(*
SPDX-FileCopyrightText: c 2026 Oleksandr Tiutyk <trofimich@gmail.com>
SPDX-License-Identifier: MIT
License: https://opensource.org/license/mit
*)

(*!
<summary>Checks the native wrapper message in HIDDEN, LOCAL and UTC modes.</summary>
<description>
Uses one task and stays at a stable address while assertions are bound to this instance.
</description>
*)

{attribute 'no_assign'}
{attribute 'no_explicit_call' := 'do not call this function block directly'}
FUNCTION_BLOCK SystemExceptionTimestampFormattingTest EXTENDS TOF_Testing.SingleCycleTest
VAR_STAT
	{attribute 'hide'}
	_ClassName : STRING := __POUNAME();
END_VAR

(*!
<summary>Checks the native wrapper message in HIDDEN, LOCAL and UTC modes.</summary>
<description>
Uses the borrowed wrapper during one callback. The timestamp expectations use the IEC conversion of
captured values and a separately assembled expected message.
</description>
*)
METHOD PROTECTED ExecuteTest
VAR
	exception : TOF_Core.IException;
	hidden : TOF_Core.ERROR_MESSAGE;
	message : TOF_Core.ERROR_MESSAGE;
	expected : WSTRING(255);
	formattingFailed : BOOL;
END_VAR
exception := TOF_Core.ExceptionManager.GetLastException(
	exceptionCode := __SYSTEM.ExceptionCode.RTSEXCPT_ACCESS_VIOLATION,
	catchPointNamespaceName := 'TimestampTest',
	catchPointPOUName := 'NativeCatch',
	catchPointPosition := 'P1'
);

IF exception = 0 THEN
	RecordFailure(message := "The captured native code must provide a wrapper");
	RETURN;
END_IF

hidden := exception.GetMessage(timestampDisplayMode := TOF_Core.TIMESTAMP_DISPLAY_MODE.HIDDEN);
Assert.ThatBool(
	actual := Tc2_Standard.WRIGHT(STR := hidden, SIZE := 31) = "TimestampTest.NativeCatch at P1",
	message := "The hidden timestamp mode must end with the supplied catch location"
).IsTrue();

expected := Tc2_Utilities.WCONCAT(STR1 := hidden, STR2 := " at ");
expected := Tc2_Utilities.WCONCAT(STR1 := expected, STR2 := TO_WSTRING(exception.LocalTimestamp));
formattingFailed := FALSE;

// A formatter exception is recorded for this mode before proceeding to the next check.
__TRY
	message := exception.GetMessage(timestampDisplayMode := TOF_Core.TIMESTAMP_DISPLAY_MODE.LOCAL);
__CATCH
	formattingFailed := TRUE;
__ENDTRY

Assert.ThatBool(
	actual := NOT formattingFailed AND_THEN message = expected,
	message := "LOCAL must append its captured timestamp"
).IsTrue();

expected := Tc2_Utilities.WCONCAT(STR1 := hidden, STR2 := " at ");
expected := Tc2_Utilities.WCONCAT(STR1 := expected, STR2 := TO_WSTRING(exception.UtcTimestamp));
expected := Tc2_Utilities.WCONCAT(STR1 := expected, STR2 := "UTC");
formattingFailed := FALSE;

// A formatter exception is recorded for this mode before proceeding to the next check.
__TRY
	message := exception.GetMessage(timestampDisplayMode := TOF_Core.TIMESTAMP_DISPLAY_MODE.UTC);
__CATCH
	formattingFailed := TRUE;
__ENDTRY

Assert.ThatBool(
	actual := NOT formattingFailed AND_THEN message = expected,
	message := "UTC must append its captured timestamp and UTC suffix"
).IsTrue();

message := exception.GetMessage(timestampDisplayMode := TOF_Core.TIMESTAMP_DISPLAY_MODE.HIDDEN);
Assert.ThatBool(
	actual := message = hidden,
	message := "Timestamp formatting must preserve the underlying diagnostic"
).IsTrue();
END_METHOD

//! <summary>Borrows the concrete class name. Callers must not modify it.</summary>
{attribute 'monitoring' := 'call'}
PROPERTY ClassName : REFERENCE TO STRING
GET
ClassName REF= _ClassName;
END_GET
END_PROPERTY

//! <summary>Borrows the compiler-initialized namespace name. Callers must not modify it.</summary>
{attribute 'monitoring' := 'call'}
PROPERTY NamespaceName : REFERENCE TO STRING
GET
NamespaceName REF= CurrentNamespace.Name;
END_GET
END_PROPERTY

//! <summary>Reports the concrete instance size in bytes.</summary>
{attribute 'monitoring' := 'call'}
PROPERTY SelfSize : ULINT
GET
SelfSize := XSIZEOF(THIS^);
END_GET
END_PROPERTY

END_FUNCTION_BLOCK

(* stored: Version 1.1.0.1
   POU SystemExceptionTimestampFormattingTest: Id {e83b71ae-bb4e-4244-9728-daa0918d9f8f}, SpecialFunc None
   Method ExecuteTest: Id {2c6ac86b-4219-41fc-a242-e028683b0364}
   Property ClassName: Id {981ad815-2bf8-4329-b7e5-a2ce87a55d1d}
   Get Get: Id {11f663e2-dcde-45ce-b8ae-111be164bd13}
   Property NamespaceName: Id {7302e617-f19e-437f-97b7-e0ac1e859d37}
   Get Get: Id {c12b7034-59b7-40c2-874f-39325b978ebe}
   Property SelfSize: Id {5f4c46b7-fe9e-4c6e-8ee0-501fd05f0108}
   Get Get: Id {5b79ecec-6691-4d47-9387-b1e75de529d1} *)
